TYPE ST_SafeIn_PlcOut :
STRUCT
	ES1_PB_Restart						:BOOL;
	ES2_PB_Restart						:BOOL;
	ES3_PB_Restart						:BOOL;
	ES4_PB_Restart						:BOOL;
	
	ES1_HMI_PB_Button						:BOOL:=TRUE;
	ES2_HMI_PB_Button						:BOOL:=TRUE;
	ES3_HMI_PB_Button						:BOOL:=TRUE;
	ES4_HMI_PB_Button						:BOOL:=TRUE;
	
END_STRUCT
END_TYPE

(* stored: Version 1.1.0.1, ProductVersion 3.1.4024.13
   DUT ST_SafeIn_PlcOut: Id {ccb37e05-6450-4451-b387-f66ff2ebdc94} *)
